(* IEC 61131-3 sources: llm-plc-st-eval/data/processed_v2_primera/gpt-4o/B6/few_shot, 3 files *)

(* ---- ejec_1.st ---- *)
FUNCTION_BLOCK FB_Baliza
VAR_INPUT
    alarma : BOOL; (* Condición de alarma *)
END_VAR
VAR_OUTPUT
    lampara : BOOL; (* Lámpara de la baliza *)
END_VAR
VAR
    tParpadeo : TON; (* Temporizador de parpadeo *)
    estadoParpadeo : BOOL; (* Estado interno de parpadeo *)
END_VAR

(* Temporizador para controlar el parpadeo de la lámpara *)
tParpadeo(IN := alarma AND NOT tParpadeo.Q, PT := T#1S);

(* Alterna el estado de la lámpara cada segundo mientras hay alarma *)
IF alarma THEN
    IF tParpadeo.Q THEN
        estadoParpadeo := NOT estadoParpadeo;
        tParpadeo(IN := FALSE); (* Reinicia el temporizador *)
    END_IF;
    lampara := estadoParpadeo;
ELSE
    lampara := FALSE; (* Lámpara apagada sin alarma *)
    estadoParpadeo := FALSE; (* Reinicia el estado de parpadeo *)
END_IF;
END_FUNCTION_BLOCK

(* ---- ejec_2.st ---- *)
FUNCTION_BLOCK FB_Baliza
VAR_INPUT
    alarma : BOOL; (* Condición de alarma *)
END_VAR
VAR_OUTPUT
    lampara : BOOL; (* Lámpara de la baliza *)
END_VAR
VAR
    tParpadeo : TON; (* Temporizador de parpadeo *)
    estadoParpadeo : BOOL; (* Estado interno de parpadeo *)
END_VAR

(* Temporizador para el parpadeo de la lámpara *)
tParpadeo(IN := alarma AND NOT tParpadeo.Q, PT := T#1S);

(* Alterna el estado de parpadeo cada segundo mientras la alarma está activa *)
IF tParpadeo.Q THEN
    estadoParpadeo := NOT estadoParpadeo;
    tParpadeo(IN := FALSE); (* Reinicia el temporizador *)
END_IF

(* La lámpara parpadea si hay alarma, de lo contrario permanece apagada *)
lampara := alarma AND estadoParpadeo;
END_FUNCTION_BLOCK

(* ---- ejec_3.st ---- *)
FUNCTION_BLOCK FB_Baliza
VAR_INPUT
    alarma : BOOL; (* Condición de alarma *)
END_VAR
VAR_OUTPUT
    lampara : BOOL; (* Lámpara de la baliza *)
END_VAR
VAR
    tParpadeo : TON; (* Temporizador de parpadeo *)
    estado : BOOL; (* Estado interno para alternar la lámpara *)
END_VAR

(* Temporizador de parpadeo de 1 segundo *)
tParpadeo(IN := alarma AND NOT tParpadeo.Q, PT := T#1S);

(* Alterna el estado de la lámpara cada segundo mientras hay alarma *)
IF tParpadeo.Q THEN
    estado := NOT estado;
    tParpadeo(IN := FALSE); (* Reinicia el temporizador *)
END_IF;

(* La lámpara parpadea si hay alarma, apagada si no hay alarma *)
lampara := alarma AND estado;
END_FUNCTION_BLOCK
